// Generated by voz_llm_plc_agent
// Target: Siemens TIA Portal V18 - SCL external source
// Review and compile before any download to physical hardware.

FUNCTION_BLOCK "PLC_PRG"
{ S7_Optimized_Access := 'TRUE' }
VERSION : 0.1
VAR_INPUT
   I_Piece_Sensor : Bool := FALSE;
   I_Emergency : Bool := FALSE;
END_VAR
VAR_OUTPUT
   Q_Aux_Output : Bool := FALSE;
END_VAR
VAR
   C_PulseCount {InstructionName := 'CTU_INT'; LibVersion := '1.0'} : CTU_INT;
   R_SensorPulse {InstructionName := 'R_TRIG'; LibVersion := '1.0'} : R_TRIG;
   M_PulseCount_Done : Bool;
   M_PulseCount_CV : Int;
END_VAR
BEGIN
(* Conteo de pulsos: CTU con salidas explicitas (alcanzado = #M_PulseCount_Done, valor = #M_PulseCount_CV) *)
#R_SensorPulse(CLK := #I_Piece_Sensor);
#C_PulseCount(CU := #R_SensorPulse.Q, R := FALSE OR #I_Emergency, PV := 5, Q => #M_PulseCount_Done, CV => #M_PulseCount_CV);
#Q_Aux_Output := #M_PulseCount_Done AND NOT #I_Emergency;
END_FUNCTION_BLOCK

DATA_BLOCK "DB_PLC_PRG"
{ S7_Optimized_Access := 'TRUE' }
VERSION : 0.1
NON_RETAIN
"PLC_PRG"
BEGIN
END_DATA_BLOCK

ORGANIZATION_BLOCK "Main"
{ S7_Optimized_Access := 'TRUE' }
VERSION : 0.1
BEGIN
   "DB_PLC_PRG"(
      I_Piece_Sensor := "I_Piece_Sensor",
      I_Emergency := "I_Emergency",
      Q_Aux_Output => "Q_Aux_Output"
   );
END_ORGANIZATION_BLOCK
